(* IEC 61131-3 sources: codesys-api/examples/mqtt_large_payload/st/bcnf_style, 5 files *)

(* ---- AppendGroupBool.st ---- *)
FUNCTION AppendGroupBool : BOOL
// Appends ", 0" or ", 1" to a BCNF-style group line, like INT_TO_STRING(BOOL_TO_INT(x)) in BCNF.
VAR_INPUT
	pBuffer : POINTER TO BYTE;
	Capacity : UDINT;
	Value : BOOL;
END_VAR
VAR_IN_OUT
	Used : UDINT;
END_VAR
// ---- implementation ----
AppendGroupBool := AppendText(pBuffer := pBuffer, Capacity := Capacity, Text := SEL(Value, ', 0', ', 1'), Used := Used);

(* ---- AppendGroupReal.st ---- *)
FUNCTION AppendGroupReal : BOOL
// Appends ", <value>" to a BCNF-style group line, rounded to two decimals exactly as
// FB_InterlockMatrix.StringPublication does. FALSE (and nothing appended) if it would not fit.
VAR_INPUT
	pBuffer : POINTER TO BYTE;
	Capacity : UDINT;
	Value : REAL;
END_VAR
VAR_IN_OUT
	Used : UDINT;
END_VAR
VAR
	Text : STRING(40);
END_VAR
// ---- implementation ----
Text := CONCAT(', ', REAL_TO_STRING(DINT_TO_REAL(TRUNC(Value * 100.0 + SEL(Value >= 0.0, -0.5, 0.5))) / 100.0));
AppendGroupReal := AppendText(pBuffer := pBuffer, Capacity := Capacity, Text := Text, Used := Used);

(* ---- AppendTagLine.st ---- *)
FUNCTION AppendTagLine : BOOL
// Appends "<Name>:<Value>\n", the line format the bridge ingests directly, without a publish map.
// All or nothing: if the whole line doesn't fit, the buffer is left as it was and FALSE is returned.
VAR_INPUT
	pBuffer : POINTER TO BYTE;
	Capacity : UDINT;
	Name : STRING(64);                  // the bridge's tag key for this value
	Value : STRING(40);                 // already formatted, e.g. by REAL_TO_STRING
END_VAR
VAR_IN_OUT
	Used : UDINT;
END_VAR
VAR
	Start : UDINT;
END_VAR
// ---- implementation ----
Start := Used;
AppendTagLine := AppendText(pBuffer := pBuffer, Capacity := Capacity, Text := Name, Used := Used)
	AND_THEN AppendText(pBuffer := pBuffer, Capacity := Capacity, Text := ':', Used := Used)
	AND_THEN AppendText(pBuffer := pBuffer, Capacity := Capacity, Text := Value, Used := Used)
	AND_THEN AppendText(pBuffer := pBuffer, Capacity := Capacity, Text := '$N', Used := Used);
IF NOT AppendTagLine AND pBuffer <> 0 THEN
	Used := Start;
	pBuffer[Start] := 0;
END_IF

(* ---- BcnfPayloadExample.st ---- *)
PROGRAM BcnfPayloadExample
// Sketch of BCNF's StringPublication without the 255-character cap: every group goes into one
// buffer, one "[GROUP, v1, v2, ...]" line per group, so a single publisher sends all of them.
// The values are copied into arrays first; that snapshot is also what a separate MQTT task needs.
// Compiled against the demo project; not run on a PLC.
VAR_INPUT
	IsBuildRequested : BOOL;            // set by the publish timer, not every scan
END_VAR
VAR_OUTPUT
	IsBuildOk : BOOL;                   // FALSE: buffer too small, do not publish this message
	PayloadLength : UDINT;
END_VAR
VAR
	Analog : ARRAY[1..14] OF REAL;      // AIT_1508_V, FIT_1506_F, ... in publish-map order
	Digital : ARRAY[1..9] OF BOOL;      // BCNF_H_E_STOP, LSL_1503_S, ...
	Payload : STRING(4000);
	Used : UDINT;
	Index : INT;
END_VAR
// ---- implementation ----
IF NOT IsBuildRequested THEN
	RETURN;   // BCNF rebuilds its strings every scan today; once per publish is enough
END_IF

// Snapshot (in BCNF: Analog[1] := AIT_1508_V; Analog[2] := FIT_1506_F; ...)

Used := 0;
Payload := '';
IsBuildOk := AppendText(pBuffer := ADR(Payload), Capacity := SIZEOF(Payload), Text := '[BCNF_ANALOG', Used := Used);
FOR Index := 1 TO 14 DO
	IsBuildOk := IsBuildOk AND_THEN AppendGroupReal(pBuffer := ADR(Payload), Capacity := SIZEOF(Payload), Value := Analog[Index], Used := Used);
END_FOR
IsBuildOk := IsBuildOk AND_THEN AppendText(pBuffer := ADR(Payload), Capacity := SIZEOF(Payload), Text := ']$N[BCNF_DIGITAL', Used := Used);
FOR Index := 1 TO 9 DO
	IsBuildOk := IsBuildOk AND_THEN AppendGroupBool(pBuffer := ADR(Payload), Capacity := SIZEOF(Payload), Value := Digital[Index], Used := Used);
END_FOR
IsBuildOk := IsBuildOk AND_THEN AppendText(pBuffer := ADR(Payload), Capacity := SIZEOF(Payload), Text := ']$N', Used := Used);
// ... the same for BCNF_ALARM, BCNF_SETPOINT_1 and _2 (one line once the bridge's publish map
// has a single setpoint entry), BCNF_OUTPUT_OTHER and BCNF_STATUS_STRING.
PayloadLength := Used;
// Publish with PayloadString := ADR(Payload) only when IsBuildOk is TRUE.

(* ---- BcnfStringPublicationCopy.st ---- *)
PROGRAM BcnfStringPublicationCopy
// BCNF's FB_InterlockMatrix.StringPublication, copied verbatim from PLC_BCNF_4_16_26.project, with the
// tags it reads declared using their BCNF types and non-zero values. Generated by
// make_bcnf_copy.py. PLC_PRG calls it every scan when IsBcnfEveryScanEnabled is TRUE,
// to measure what rebuilding BCNF's payload strings every scan costs. Its BuildTagValue action
// builds the same values in the bridge's tag:value line format instead.
VAR
	BCNF_ANALOG_STRING : STRING(255);
	AIT_1508_V : REAL := 16.88;
	FIT_1506_F : REAL := 30.59;
	FIT_1520_F : REAL := 44.30;
	PT_1513_P : REAL := 58.01;
	PT_1516_P : REAL := 71.72;
	QIT_1507_V : REAL := 85.43;
	QIT_1518_V : REAL := 99.14;
	REC_1525_V : REAL := 112.85;
	REJ_1526_V : REAL := 126.56;
	TT_1509_T : REAL := 140.27;
	VFD_1512C_V : REAL := 153.98;
	VFD_1512F_V : REAL := 167.69;
	VFD_1512T_V : REAL := 181.40;
	VFD_1512V_V : REAL := 195.11;
	BCNF_DIGITAL_STRING : STRING(255);
	BCNF_H_E_STOP : BOOL;
	LSL_1503_S : BOOL;
	LSS_E_STOP : BOOL := TRUE;
	LS_1521_S : BOOL;
	LS_1522_S : BOOL;
	LS_1523_S : BOOL := TRUE;
	LS_1524_S : BOOL;
	P_1502FB : BOOL;
	P_1504 : BOOL := TRUE;
	BCNF_ALARM_STRING : STRING(255);
	AIT_1508H : BOOL;
	AIT_1508HH : BOOL;
	AIT_1508L : BOOL := TRUE;
	AIT_1508LL : BOOL;
	BCNF_E_STOP : BOOL;
	BCNF_E_STOPH : BOOL := TRUE;
	BCNF_H_E_STOPH : BOOL;
	CONC_BCNF_PLC_STATUSH : BOOL;
	FIT_1506H : BOOL := TRUE;
	FIT_1506HH : BOOL;
	FIT_1520H : BOOL;
	FIT_1520HH : BOOL := TRUE;
	LSL_1503LL : BOOL;
	LSS_E_STOPH : BOOL;
	LS_1521LL : BOOL := TRUE;
	LS_1522L : BOOL;
	LS_1523H : BOOL;
	LS_1524HH : BOOL := TRUE;
	PT_1513H : BOOL;
	PT_1513HH : BOOL;
	PT_1513L : BOOL := TRUE;
	PT_1513LL : BOOL;
	PT_1516H : BOOL;
	PT_1516HH : BOOL := TRUE;
	PT_1516L : BOOL;
	PT_1516LL : BOOL;
	P_1502FBHH : BOOL := TRUE;
	QIT_1507H : BOOL;
	QIT_1507HH : BOOL;
	QIT_1518H : BOOL := TRUE;
	QIT_1518HH : BOOL;
	TT_1509H : BOOL;
	TT_1509HH : BOOL := TRUE;
	TT_1509L : BOOL;
	TT_1509LL : BOOL;
	VFD_1512CH : BOOL := TRUE;
	VFD_1512CHH : BOOL;
	VFD_1512FH : BOOL;
	VFD_1512FHH : BOOL := TRUE;
	VFD_1512TH : BOOL;
	VFD_1512THH : BOOL;
	VFD_1512VH : BOOL := TRUE;
	VFD_1512VHH : BOOL;
	BCNF_SETPOINT_STRING_1 : STRING(255);
	AIT_1508_HH_SP : REAL := 208.82;
	AIT_1508_H_SP : REAL := 222.53;
	AIT_1508_LL_SP : REAL := 236.24;
	AIT_1508_L_SP : REAL := 249.95;
	FIT_1506_HH_SP : REAL := 263.66;
	FIT_1506_H_SP : REAL := 277.37;
	FIT_1520_HH_SP : REAL := 291.08;
	FIT_1520_H_SP : REAL := 304.79;
	PT_1513_HH_SP : REAL := 318.50;
	PT_1513_H_SP : REAL := 332.21;
	PT_1513_LL_SP : REAL := 345.92;
	PT_1513_L_SP : REAL := 359.63;
	PT_1516_HH_SP : REAL := 373.34;
	PT_1516_H_SP : REAL := 387.05;
	PT_1516_LL_SP : REAL := 400.76;
	PT_1516_L_SP : REAL := 414.47;
	QIT_1507_HH_SP : REAL := 428.18;
	QIT_1507_H_SP : REAL := 441.89;
	QIT_1518_HH_SP : REAL := 455.60;
	QIT_1518_H_SP : REAL := 469.31;
	TT_1509_HH_SP : REAL := 483.02;
	TT_1509_H_SP : REAL := 496.73;
	TT_1509_LL_SP : REAL := 510.44;
	TT_1509_L_SP : REAL := 524.15;
	VFD_1512C_HH_SP : REAL := 537.86;
	VFD_1512C_H_SP : REAL := 551.57;
	BCNF_SETPOINT_STRING_2 : STRING(255);
	VFD_1512F_HH_SP : REAL := 565.28;
	VFD_1512F_H_SP : REAL := 578.99;
	VFD_1512T_HH_SP : REAL := 592.70;
	VFD_1512T_H_SP : REAL := 606.41;
	VFD_1512V_HH_SP : REAL := 620.12;
	VFD_1512V_H_SP : REAL := 633.83;
	BCNF_OUTPUT_OTHER_STRING : STRING(255);
	P_1502_OUTPUT : BOOL;
	VFD_1512FSP : REAL := 647.54;
	VFD_1512SP : REAL := 661.25;
	BCNF_STATUS_STRING : STRING(255);
	Heartbeat : DINT := 18234;
	CONC_BCNF_PLC_STATUS : BOOL := TRUE;
	fullPayload_BCNF_ANALOG_STRING : STRING(255);
	fullPayload_BCNF_DIGITAL_STRING : STRING(255);
	fullPayload_BCNF_ALARM_STRING : STRING(255);
	fullPayload_BCNF_SETPOINT_STRING_1 : STRING(255);
	fullPayload_BCNF_SETPOINT_STRING_2 : STRING(255);
	fullPayload_BCNF_OUTPUT_OTHER_STRING : STRING(255);
	fullPayload_BCNF_STATUS_STRING : STRING(255);
	// BuildTagValue action: the same values as one tag:value line each
	TagValuePayload : STRING(4000);
	TagValueUsed : UDINT;
	IsTagValueBuildOk : BOOL;
END_VAR
// ---- implementation ----
// ===== DATA PUBLICATION STRING BUILDING =====
// This code should be placed in a StringPublication action

// Build BCNF_ANALOG string
BCNF_ANALOG_STRING := '[BCNF_ANALOG, ';
BCNF_ANALOG_STRING := CONCAT(BCNF_ANALOG_STRING, REAL_TO_STRING(DINT_TO_REAL(TRUNC(AIT_1508_V * 100.0 + SEL(AIT_1508_V >= 0.0, -0.5, 0.5))) / 100.0));
BCNF_ANALOG_STRING := CONCAT(BCNF_ANALOG_STRING, ', ');
BCNF_ANALOG_STRING := CONCAT(BCNF_ANALOG_STRING, REAL_TO_STRING(DINT_TO_REAL(TRUNC(FIT_1506_F * 100.0 + SEL(FIT_1506_F >= 0.0, -0.5, 0.5))) / 100.0));
BCNF_ANALOG_STRING := CONCAT(BCNF_ANALOG_STRING, ', ');
BCNF_ANALOG_STRING := CONCAT(BCNF_ANALOG_STRING, REAL_TO_STRING(DINT_TO_REAL(TRUNC(FIT_1520_F * 100.0 + SEL(FIT_1520_F >= 0.0, -0.5, 0.5))) / 100.0));
BCNF_ANALOG_STRING := CONCAT(BCNF_ANALOG_STRING, ', ');
BCNF_ANALOG_STRING := CONCAT(BCNF_ANALOG_STRING, REAL_TO_STRING(DINT_TO_REAL(TRUNC(PT_1513_P * 100.0 + SEL(PT_1513_P >= 0.0, -0.5, 0.5))) / 100.0));
BCNF_ANALOG_STRING := CONCAT(BCNF_ANALOG_STRING, ', ');
BCNF_ANALOG_STRING := CONCAT(BCNF_ANALOG_STRING, REAL_TO_STRING(DINT_TO_REAL(TRUNC(PT_1516_P * 100.0 + SEL(PT_1516_P >= 0.0, -0.5, 0.5))) / 100.0));
BCNF_ANALOG_STRING := CONCAT(BCNF_ANALOG_STRING, ', ');
BCNF_ANALOG_STRING := CONCAT(BCNF_ANALOG_STRING, REAL_TO_STRING(DINT_TO_REAL(TRUNC(QIT_1507_V * 100.0 + SEL(QIT_1507_V >= 0.0, -0.5, 0.5))) / 100.0));
BCNF_ANALOG_STRING := CONCAT(BCNF_ANALOG_STRING, ', ');
BCNF_ANALOG_STRING := CONCAT(BCNF_ANALOG_STRING, REAL_TO_STRING(DINT_TO_REAL(TRUNC(QIT_1518_V * 100.0 + SEL(QIT_1518_V >= 0.0, -0.5, 0.5))) / 100.0));
BCNF_ANALOG_STRING := CONCAT(BCNF_ANALOG_STRING, ', ');
BCNF_ANALOG_STRING := CONCAT(BCNF_ANALOG_STRING, REAL_TO_STRING(DINT_TO_REAL(TRUNC(REC_1525_V * 100.0 + SEL(REC_1525_V >= 0.0, -0.5, 0.5))) / 100.0));
BCNF_ANALOG_STRING := CONCAT(BCNF_ANALOG_STRING, ', ');
BCNF_ANALOG_STRING := CONCAT(BCNF_ANALOG_STRING, REAL_TO_STRING(DINT_TO_REAL(TRUNC(REJ_1526_V * 100.0 + SEL(REJ_1526_V >= 0.0, -0.5, 0.5))) / 100.0));
BCNF_ANALOG_STRING := CONCAT(BCNF_ANALOG_STRING, ', ');
BCNF_ANALOG_STRING := CONCAT(BCNF_ANALOG_STRING, REAL_TO_STRING(DINT_TO_REAL(TRUNC(TT_1509_T * 100.0 + SEL(TT_1509_T >= 0.0, -0.5, 0.5))) / 100.0));
BCNF_ANALOG_STRING := CONCAT(BCNF_ANALOG_STRING, ', ');
BCNF_ANALOG_STRING := CONCAT(BCNF_ANALOG_STRING, REAL_TO_STRING(DINT_TO_REAL(TRUNC(VFD_1512C_V * 100.0 + SEL(VFD_1512C_V >= 0.0, -0.5, 0.5))) / 100.0));
BCNF_ANALOG_STRING := CONCAT(BCNF_ANALOG_STRING, ', ');
BCNF_ANALOG_STRING := CONCAT(BCNF_ANALOG_STRING, REAL_TO_STRING(DINT_TO_REAL(TRUNC(VFD_1512F_V * 100.0 + SEL(VFD_1512F_V >= 0.0, -0.5, 0.5))) / 100.0));
BCNF_ANALOG_STRING := CONCAT(BCNF_ANALOG_STRING, ', ');
BCNF_ANALOG_STRING := CONCAT(BCNF_ANALOG_STRING, REAL_TO_STRING(DINT_TO_REAL(TRUNC(VFD_1512T_V * 100.0 + SEL(VFD_1512T_V >= 0.0, -0.5, 0.5))) / 100.0));
BCNF_ANALOG_STRING := CONCAT(BCNF_ANALOG_STRING, ', ');
BCNF_ANALOG_STRING := CONCAT(BCNF_ANALOG_STRING, REAL_TO_STRING(DINT_TO_REAL(TRUNC(VFD_1512V_V * 100.0 + SEL(VFD_1512V_V >= 0.0, -0.5, 0.5))) / 100.0));
BCNF_ANALOG_STRING := CONCAT(BCNF_ANALOG_STRING, ']');

// Build BCNF_DIGITAL string
BCNF_DIGITAL_STRING := '[BCNF_DIGITAL, ';
BCNF_DIGITAL_STRING := CONCAT(BCNF_DIGITAL_STRING, INT_TO_STRING(BOOL_TO_INT(BCNF_H_E_STOP)));
BCNF_DIGITAL_STRING := CONCAT(BCNF_DIGITAL_STRING, ', ');
BCNF_DIGITAL_STRING := CONCAT(BCNF_DIGITAL_STRING, INT_TO_STRING(BOOL_TO_INT(LSL_1503_S)));
BCNF_DIGITAL_STRING := CONCAT(BCNF_DIGITAL_STRING, ', ');
BCNF_DIGITAL_STRING := CONCAT(BCNF_DIGITAL_STRING, INT_TO_STRING(BOOL_TO_INT(LSS_E_STOP)));
BCNF_DIGITAL_STRING := CONCAT(BCNF_DIGITAL_STRING, ', ');
BCNF_DIGITAL_STRING := CONCAT(BCNF_DIGITAL_STRING, INT_TO_STRING(BOOL_TO_INT(LS_1521_S)));
BCNF_DIGITAL_STRING := CONCAT(BCNF_DIGITAL_STRING, ', ');
BCNF_DIGITAL_STRING := CONCAT(BCNF_DIGITAL_STRING, INT_TO_STRING(BOOL_TO_INT(LS_1522_S)));
BCNF_DIGITAL_STRING := CONCAT(BCNF_DIGITAL_STRING, ', ');
BCNF_DIGITAL_STRING := CONCAT(BCNF_DIGITAL_STRING, INT_TO_STRING(BOOL_TO_INT(LS_1523_S)));
BCNF_DIGITAL_STRING := CONCAT(BCNF_DIGITAL_STRING, ', ');
BCNF_DIGITAL_STRING := CONCAT(BCNF_DIGITAL_STRING, INT_TO_STRING(BOOL_TO_INT(LS_1524_S)));
BCNF_DIGITAL_STRING := CONCAT(BCNF_DIGITAL_STRING, ', ');
BCNF_DIGITAL_STRING := CONCAT(BCNF_DIGITAL_STRING, INT_TO_STRING(BOOL_TO_INT(P_1502FB)));
BCNF_DIGITAL_STRING := CONCAT(BCNF_DIGITAL_STRING, ', ');
BCNF_DIGITAL_STRING := CONCAT(BCNF_DIGITAL_STRING, INT_TO_STRING(BOOL_TO_INT(P_1504)));
BCNF_DIGITAL_STRING := CONCAT(BCNF_DIGITAL_STRING, ']');

// Build BCNF_ALARM string
BCNF_ALARM_STRING := '[BCNF_ALARM, ';
BCNF_ALARM_STRING := CONCAT(BCNF_ALARM_STRING, INT_TO_STRING(BOOL_TO_INT(AIT_1508H)));
BCNF_ALARM_STRING := CONCAT(BCNF_ALARM_STRING, ', ');
BCNF_ALARM_STRING := CONCAT(BCNF_ALARM_STRING, INT_TO_STRING(BOOL_TO_INT(AIT_1508HH)));
BCNF_ALARM_STRING := CONCAT(BCNF_ALARM_STRING, ', ');
BCNF_ALARM_STRING := CONCAT(BCNF_ALARM_STRING, INT_TO_STRING(BOOL_TO_INT(AIT_1508L)));
BCNF_ALARM_STRING := CONCAT(BCNF_ALARM_STRING, ', ');
BCNF_ALARM_STRING := CONCAT(BCNF_ALARM_STRING, INT_TO_STRING(BOOL_TO_INT(AIT_1508LL)));
BCNF_ALARM_STRING := CONCAT(BCNF_ALARM_STRING, ', ');
BCNF_ALARM_STRING := CONCAT(BCNF_ALARM_STRING, INT_TO_STRING(BOOL_TO_INT(BCNF_E_STOP)));
BCNF_ALARM_STRING := CONCAT(BCNF_ALARM_STRING, ', ');
BCNF_ALARM_STRING := CONCAT(BCNF_ALARM_STRING, INT_TO_STRING(BOOL_TO_INT(BCNF_E_STOPH)));
BCNF_ALARM_STRING := CONCAT(BCNF_ALARM_STRING, ', ');
BCNF_ALARM_STRING := CONCAT(BCNF_ALARM_STRING, INT_TO_STRING(BOOL_TO_INT(BCNF_H_E_STOPH)));
BCNF_ALARM_STRING := CONCAT(BCNF_ALARM_STRING, ', ');
BCNF_ALARM_STRING := CONCAT(BCNF_ALARM_STRING, INT_TO_STRING(BOOL_TO_INT(CONC_BCNF_PLC_STATUSH)));
BCNF_ALARM_STRING := CONCAT(BCNF_ALARM_STRING, ', ');
BCNF_ALARM_STRING := CONCAT(BCNF_ALARM_STRING, INT_TO_STRING(BOOL_TO_INT(FIT_1506H)));
BCNF_ALARM_STRING := CONCAT(BCNF_ALARM_STRING, ', ');
BCNF_ALARM_STRING := CONCAT(BCNF_ALARM_STRING, INT_TO_STRING(BOOL_TO_INT(FIT_1506HH)));
BCNF_ALARM_STRING := CONCAT(BCNF_ALARM_STRING, ', ');
BCNF_ALARM_STRING := CONCAT(BCNF_ALARM_STRING, INT_TO_STRING(BOOL_TO_INT(FIT_1520H)));
BCNF_ALARM_STRING := CONCAT(BCNF_ALARM_STRING, ', ');
BCNF_ALARM_STRING := CONCAT(BCNF_ALARM_STRING, INT_TO_STRING(BOOL_TO_INT(FIT_1520HH)));
BCNF_ALARM_STRING := CONCAT(BCNF_ALARM_STRING, ', ');
BCNF_ALARM_STRING := CONCAT(BCNF_ALARM_STRING, INT_TO_STRING(BOOL_TO_INT(LSL_1503LL)));
BCNF_ALARM_STRING := CONCAT(BCNF_ALARM_STRING, ', ');
BCNF_ALARM_STRING := CONCAT(BCNF_ALARM_STRING, INT_TO_STRING(BOOL_TO_INT(LSS_E_STOPH)));
BCNF_ALARM_STRING := CONCAT(BCNF_ALARM_STRING, ', ');
BCNF_ALARM_STRING := CONCAT(BCNF_ALARM_STRING, INT_TO_STRING(BOOL_TO_INT(LS_1521LL)));
BCNF_ALARM_STRING := CONCAT(BCNF_ALARM_STRING, ', ');
BCNF_ALARM_STRING := CONCAT(BCNF_ALARM_STRING, INT_TO_STRING(BOOL_TO_INT(LS_1522L)));
BCNF_ALARM_STRING := CONCAT(BCNF_ALARM_STRING, ', ');
BCNF_ALARM_STRING := CONCAT(BCNF_ALARM_STRING, INT_TO_STRING(BOOL_TO_INT(LS_1523H)));
BCNF_ALARM_STRING := CONCAT(BCNF_ALARM_STRING, ', ');
BCNF_ALARM_STRING := CONCAT(BCNF_ALARM_STRING, INT_TO_STRING(BOOL_TO_INT(LS_1524HH)));
BCNF_ALARM_STRING := CONCAT(BCNF_ALARM_STRING, ', ');
BCNF_ALARM_STRING := CONCAT(BCNF_ALARM_STRING, INT_TO_STRING(BOOL_TO_INT(PT_1513H)));
BCNF_ALARM_STRING := CONCAT(BCNF_ALARM_STRING, ', ');
BCNF_ALARM_STRING := CONCAT(BCNF_ALARM_STRING, INT_TO_STRING(BOOL_TO_INT(PT_1513HH)));
BCNF_ALARM_STRING := CONCAT(BCNF_ALARM_STRING, ', ');
BCNF_ALARM_STRING := CONCAT(BCNF_ALARM_STRING, INT_TO_STRING(BOOL_TO_INT(PT_1513L)));
BCNF_ALARM_STRING := CONCAT(BCNF_ALARM_STRING, ', ');
BCNF_ALARM_STRING := CONCAT(BCNF_ALARM_STRING, INT_TO_STRING(BOOL_TO_INT(PT_1513LL)));
BCNF_ALARM_STRING := CONCAT(BCNF_ALARM_STRING, ', ');
BCNF_ALARM_STRING := CONCAT(BCNF_ALARM_STRING, INT_TO_STRING(BOOL_TO_INT(PT_1516H)));
BCNF_ALARM_STRING := CONCAT(BCNF_ALARM_STRING, ', ');
BCNF_ALARM_STRING := CONCAT(BCNF_ALARM_STRING, INT_TO_STRING(BOOL_TO_INT(PT_1516HH)));
BCNF_ALARM_STRING := CONCAT(BCNF_ALARM_STRING, ', ');
BCNF_ALARM_STRING := CONCAT(BCNF_ALARM_STRING, INT_TO_STRING(BOOL_TO_INT(PT_1516L)));
BCNF_ALARM_STRING := CONCAT(BCNF_ALARM_STRING, ', ');
BCNF_ALARM_STRING := CONCAT(BCNF_ALARM_STRING, INT_TO_STRING(BOOL_TO_INT(PT_1516LL)));
BCNF_ALARM_STRING := CONCAT(BCNF_ALARM_STRING, ', ');
BCNF_ALARM_STRING := CONCAT(BCNF_ALARM_STRING, INT_TO_STRING(BOOL_TO_INT(P_1502FBHH)));
BCNF_ALARM_STRING := CONCAT(BCNF_ALARM_STRING, ', ');
BCNF_ALARM_STRING := CONCAT(BCNF_ALARM_STRING, INT_TO_STRING(BOOL_TO_INT(QIT_1507H)));
BCNF_ALARM_STRING := CONCAT(BCNF_ALARM_STRING, ', ');
BCNF_ALARM_STRING := CONCAT(BCNF_ALARM_STRING, INT_TO_STRING(BOOL_TO_INT(QIT_1507HH)));
BCNF_ALARM_STRING := CONCAT(BCNF_ALARM_STRING, ', ');
BCNF_ALARM_STRING := CONCAT(BCNF_ALARM_STRING, INT_TO_STRING(BOOL_TO_INT(QIT_1518H)));
BCNF_ALARM_STRING := CONCAT(BCNF_ALARM_STRING, ', ');
BCNF_ALARM_STRING := CONCAT(BCNF_ALARM_STRING, INT_TO_STRING(BOOL_TO_INT(QIT_1518HH)));
BCNF_ALARM_STRING := CONCAT(BCNF_ALARM_STRING, ', ');
BCNF_ALARM_STRING := CONCAT(BCNF_ALARM_STRING, INT_TO_STRING(BOOL_TO_INT(TT_1509H)));
BCNF_ALARM_STRING := CONCAT(BCNF_ALARM_STRING, ', ');
BCNF_ALARM_STRING := CONCAT(BCNF_ALARM_STRING, INT_TO_STRING(BOOL_TO_INT(TT_1509HH)));
BCNF_ALARM_STRING := CONCAT(BCNF_ALARM_STRING, ', ');
BCNF_ALARM_STRING := CONCAT(BCNF_ALARM_STRING, INT_TO_STRING(BOOL_TO_INT(TT_1509L)));
BCNF_ALARM_STRING := CONCAT(BCNF_ALARM_STRING, ', ');
BCNF_ALARM_STRING := CONCAT(BCNF_ALARM_STRING, INT_TO_STRING(BOOL_TO_INT(TT_1509LL)));
BCNF_ALARM_STRING := CONCAT(BCNF_ALARM_STRING, ', ');
BCNF_ALARM_STRING := CONCAT(BCNF_ALARM_STRING, INT_TO_STRING(BOOL_TO_INT(VFD_1512CH)));
BCNF_ALARM_STRING := CONCAT(BCNF_ALARM_STRING, ', ');
BCNF_ALARM_STRING := CONCAT(BCNF_ALARM_STRING, INT_TO_STRING(BOOL_TO_INT(VFD_1512CHH)));
BCNF_ALARM_STRING := CONCAT(BCNF_ALARM_STRING, ', ');
BCNF_ALARM_STRING := CONCAT(BCNF_ALARM_STRING, INT_TO_STRING(BOOL_TO_INT(VFD_1512FH)));
BCNF_ALARM_STRING := CONCAT(BCNF_ALARM_STRING, ', ');
BCNF_ALARM_STRING := CONCAT(BCNF_ALARM_STRING, INT_TO_STRING(BOOL_TO_INT(VFD_1512FHH)));
BCNF_ALARM_STRING := CONCAT(BCNF_ALARM_STRING, ', ');
BCNF_ALARM_STRING := CONCAT(BCNF_ALARM_STRING, INT_TO_STRING(BOOL_TO_INT(VFD_1512TH)));
BCNF_ALARM_STRING := CONCAT(BCNF_ALARM_STRING, ', ');
BCNF_ALARM_STRING := CONCAT(BCNF_ALARM_STRING, INT_TO_STRING(BOOL_TO_INT(VFD_1512THH)));
BCNF_ALARM_STRING := CONCAT(BCNF_ALARM_STRING, ', ');
BCNF_ALARM_STRING := CONCAT(BCNF_ALARM_STRING, INT_TO_STRING(BOOL_TO_INT(VFD_1512VH)));
BCNF_ALARM_STRING := CONCAT(BCNF_ALARM_STRING, ', ');
BCNF_ALARM_STRING := CONCAT(BCNF_ALARM_STRING, INT_TO_STRING(BOOL_TO_INT(VFD_1512VHH)));
BCNF_ALARM_STRING := CONCAT(BCNF_ALARM_STRING, ']');

// Build BCNF_SETPOINT string part 1
BCNF_SETPOINT_STRING_1 := '[BCNF_SETPOINT_1, ';
BCNF_SETPOINT_STRING_1 := CONCAT(BCNF_SETPOINT_STRING_1, REAL_TO_STRING(DINT_TO_REAL(TRUNC(AIT_1508_HH_SP * 100.0 + SEL(AIT_1508_HH_SP >= 0.0, -0.5, 0.5))) / 100.0));
BCNF_SETPOINT_STRING_1 := CONCAT(BCNF_SETPOINT_STRING_1, ', ');
BCNF_SETPOINT_STRING_1 := CONCAT(BCNF_SETPOINT_STRING_1, REAL_TO_STRING(DINT_TO_REAL(TRUNC(AIT_1508_H_SP * 100.0 + SEL(AIT_1508_H_SP >= 0.0, -0.5, 0.5))) / 100.0));
BCNF_SETPOINT_STRING_1 := CONCAT(BCNF_SETPOINT_STRING_1, ', ');
BCNF_SETPOINT_STRING_1 := CONCAT(BCNF_SETPOINT_STRING_1, REAL_TO_STRING(DINT_TO_REAL(TRUNC(AIT_1508_LL_SP * 100.0 + SEL(AIT_1508_LL_SP >= 0.0, -0.5, 0.5))) / 100.0));
BCNF_SETPOINT_STRING_1 := CONCAT(BCNF_SETPOINT_STRING_1, ', ');
BCNF_SETPOINT_STRING_1 := CONCAT(BCNF_SETPOINT_STRING_1, REAL_TO_STRING(DINT_TO_REAL(TRUNC(AIT_1508_L_SP * 100.0 + SEL(AIT_1508_L_SP >= 0.0, -0.5, 0.5))) / 100.0));
BCNF_SETPOINT_STRING_1 := CONCAT(BCNF_SETPOINT_STRING_1, ', ');
BCNF_SETPOINT_STRING_1 := CONCAT(BCNF_SETPOINT_STRING_1, REAL_TO_STRING(DINT_TO_REAL(TRUNC(FIT_1506_HH_SP * 100.0 + SEL(FIT_1506_HH_SP >= 0.0, -0.5, 0.5))) / 100.0));
BCNF_SETPOINT_STRING_1 := CONCAT(BCNF_SETPOINT_STRING_1, ', ');
BCNF_SETPOINT_STRING_1 := CONCAT(BCNF_SETPOINT_STRING_1, REAL_TO_STRING(DINT_TO_REAL(TRUNC(FIT_1506_H_SP * 100.0 + SEL(FIT_1506_H_SP >= 0.0, -0.5, 0.5))) / 100.0));
BCNF_SETPOINT_STRING_1 := CONCAT(BCNF_SETPOINT_STRING_1, ', ');
BCNF_SETPOINT_STRING_1 := CONCAT(BCNF_SETPOINT_STRING_1, REAL_TO_STRING(DINT_TO_REAL(TRUNC(FIT_1520_HH_SP * 100.0 + SEL(FIT_1520_HH_SP >= 0.0, -0.5, 0.5))) / 100.0));
BCNF_SETPOINT_STRING_1 := CONCAT(BCNF_SETPOINT_STRING_1, ', ');
BCNF_SETPOINT_STRING_1 := CONCAT(BCNF_SETPOINT_STRING_1, REAL_TO_STRING(DINT_TO_REAL(TRUNC(FIT_1520_H_SP * 100.0 + SEL(FIT_1520_H_SP >= 0.0, -0.5, 0.5))) / 100.0));
BCNF_SETPOINT_STRING_1 := CONCAT(BCNF_SETPOINT_STRING_1, ', ');
BCNF_SETPOINT_STRING_1 := CONCAT(BCNF_SETPOINT_STRING_1, REAL_TO_STRING(DINT_TO_REAL(TRUNC(PT_1513_HH_SP * 100.0 + SEL(PT_1513_HH_SP >= 0.0, -0.5, 0.5))) / 100.0));
BCNF_SETPOINT_STRING_1 := CONCAT(BCNF_SETPOINT_STRING_1, ', ');
BCNF_SETPOINT_STRING_1 := CONCAT(BCNF_SETPOINT_STRING_1, REAL_TO_STRING(DINT_TO_REAL(TRUNC(PT_1513_H_SP * 100.0 + SEL(PT_1513_H_SP >= 0.0, -0.5, 0.5))) / 100.0));
BCNF_SETPOINT_STRING_1 := CONCAT(BCNF_SETPOINT_STRING_1, ', ');
BCNF_SETPOINT_STRING_1 := CONCAT(BCNF_SETPOINT_STRING_1, REAL_TO_STRING(DINT_TO_REAL(TRUNC(PT_1513_LL_SP * 100.0 + SEL(PT_1513_LL_SP >= 0.0, -0.5, 0.5))) / 100.0));
BCNF_SETPOINT_STRING_1 := CONCAT(BCNF_SETPOINT_STRING_1, ', ');
BCNF_SETPOINT_STRING_1 := CONCAT(BCNF_SETPOINT_STRING_1, REAL_TO_STRING(DINT_TO_REAL(TRUNC(PT_1513_L_SP * 100.0 + SEL(PT_1513_L_SP >= 0.0, -0.5, 0.5))) / 100.0));
BCNF_SETPOINT_STRING_1 := CONCAT(BCNF_SETPOINT_STRING_1, ', ');
BCNF_SETPOINT_STRING_1 := CONCAT(BCNF_SETPOINT_STRING_1, REAL_TO_STRING(DINT_TO_REAL(TRUNC(PT_1516_HH_SP * 100.0 + SEL(PT_1516_HH_SP >= 0.0, -0.5, 0.5))) / 100.0));
BCNF_SETPOINT_STRING_1 := CONCAT(BCNF_SETPOINT_STRING_1, ', ');
BCNF_SETPOINT_STRING_1 := CONCAT(BCNF_SETPOINT_STRING_1, REAL_TO_STRING(DINT_TO_REAL(TRUNC(PT_1516_H_SP * 100.0 + SEL(PT_1516_H_SP >= 0.0, -0.5, 0.5))) / 100.0));
BCNF_SETPOINT_STRING_1 := CONCAT(BCNF_SETPOINT_STRING_1, ', ');
BCNF_SETPOINT_STRING_1 := CONCAT(BCNF_SETPOINT_STRING_1, REAL_TO_STRING(DINT_TO_REAL(TRUNC(PT_1516_LL_SP * 100.0 + SEL(PT_1516_LL_SP >= 0.0, -0.5, 0.5))) / 100.0));
BCNF_SETPOINT_STRING_1 := CONCAT(BCNF_SETPOINT_STRING_1, ', ');
BCNF_SETPOINT_STRING_1 := CONCAT(BCNF_SETPOINT_STRING_1, REAL_TO_STRING(DINT_TO_REAL(TRUNC(PT_1516_L_SP * 100.0 + SEL(PT_1516_L_SP >= 0.0, -0.5, 0.5))) / 100.0));
BCNF_SETPOINT_STRING_1 := CONCAT(BCNF_SETPOINT_STRING_1, ', ');
BCNF_SETPOINT_STRING_1 := CONCAT(BCNF_SETPOINT_STRING_1, REAL_TO_STRING(DINT_TO_REAL(TRUNC(QIT_1507_HH_SP * 100.0 + SEL(QIT_1507_HH_SP >= 0.0, -0.5, 0.5))) / 100.0));
BCNF_SETPOINT_STRING_1 := CONCAT(BCNF_SETPOINT_STRING_1, ', ');
BCNF_SETPOINT_STRING_1 := CONCAT(BCNF_SETPOINT_STRING_1, REAL_TO_STRING(DINT_TO_REAL(TRUNC(QIT_1507_H_SP * 100.0 + SEL(QIT_1507_H_SP >= 0.0, -0.5, 0.5))) / 100.0));
BCNF_SETPOINT_STRING_1 := CONCAT(BCNF_SETPOINT_STRING_1, ', ');
BCNF_SETPOINT_STRING_1 := CONCAT(BCNF_SETPOINT_STRING_1, REAL_TO_STRING(DINT_TO_REAL(TRUNC(QIT_1518_HH_SP * 100.0 + SEL(QIT_1518_HH_SP >= 0.0, -0.5, 0.5))) / 100.0));
BCNF_SETPOINT_STRING_1 := CONCAT(BCNF_SETPOINT_STRING_1, ', ');
BCNF_SETPOINT_STRING_1 := CONCAT(BCNF_SETPOINT_STRING_1, REAL_TO_STRING(DINT_TO_REAL(TRUNC(QIT_1518_H_SP * 100.0 + SEL(QIT_1518_H_SP >= 0.0, -0.5, 0.5))) / 100.0));
BCNF_SETPOINT_STRING_1 := CONCAT(BCNF_SETPOINT_STRING_1, ', ');
BCNF_SETPOINT_STRING_1 := CONCAT(BCNF_SETPOINT_STRING_1, REAL_TO_STRING(DINT_TO_REAL(TRUNC(TT_1509_HH_SP * 100.0 + SEL(TT_1509_HH_SP >= 0.0, -0.5, 0.5))) / 100.0));
BCNF_SETPOINT_STRING_1 := CONCAT(BCNF_SETPOINT_STRING_1, ', ');
BCNF_SETPOINT_STRING_1 := CONCAT(BCNF_SETPOINT_STRING_1, REAL_TO_STRING(DINT_TO_REAL(TRUNC(TT_1509_H_SP * 100.0 + SEL(TT_1509_H_SP >= 0.0, -0.5, 0.5))) / 100.0));
BCNF_SETPOINT_STRING_1 := CONCAT(BCNF_SETPOINT_STRING_1, ', ');
BCNF_SETPOINT_STRING_1 := CONCAT(BCNF_SETPOINT_STRING_1, REAL_TO_STRING(DINT_TO_REAL(TRUNC(TT_1509_LL_SP * 100.0 + SEL(TT_1509_LL_SP >= 0.0, -0.5, 0.5))) / 100.0));
BCNF_SETPOINT_STRING_1 := CONCAT(BCNF_SETPOINT_STRING_1, ', ');
BCNF_SETPOINT_STRING_1 := CONCAT(BCNF_SETPOINT_STRING_1, REAL_TO_STRING(DINT_TO_REAL(TRUNC(TT_1509_L_SP * 100.0 + SEL(TT_1509_L_SP >= 0.0, -0.5, 0.5))) / 100.0));
BCNF_SETPOINT_STRING_1 := CONCAT(BCNF_SETPOINT_STRING_1, ', ');
BCNF_SETPOINT_STRING_1 := CONCAT(BCNF_SETPOINT_STRING_1, REAL_TO_STRING(DINT_TO_REAL(TRUNC(VFD_1512C_HH_SP * 100.0 + SEL(VFD_1512C_HH_SP >= 0.0, -0.5, 0.5))) / 100.0));
BCNF_SETPOINT_STRING_1 := CONCAT(BCNF_SETPOINT_STRING_1, ', ');
BCNF_SETPOINT_STRING_1 := CONCAT(BCNF_SETPOINT_STRING_1, REAL_TO_STRING(DINT_TO_REAL(TRUNC(VFD_1512C_H_SP * 100.0 + SEL(VFD_1512C_H_SP >= 0.0, -0.5, 0.5))) / 100.0));
BCNF_SETPOINT_STRING_1 := CONCAT(BCNF_SETPOINT_STRING_1, ']');
// Build BCNF_SETPOINT string part 2
BCNF_SETPOINT_STRING_2 := '[BCNF_SETPOINT_2, ';
BCNF_SETPOINT_STRING_2 := CONCAT(BCNF_SETPOINT_STRING_2, REAL_TO_STRING(DINT_TO_REAL(TRUNC(VFD_1512F_HH_SP * 100.0 + SEL(VFD_1512F_HH_SP >= 0.0, -0.5, 0.5))) / 100.0));
BCNF_SETPOINT_STRING_2 := CONCAT(BCNF_SETPOINT_STRING_2, ', ');
BCNF_SETPOINT_STRING_2 := CONCAT(BCNF_SETPOINT_STRING_2, REAL_TO_STRING(DINT_TO_REAL(TRUNC(VFD_1512F_H_SP * 100.0 + SEL(VFD_1512F_H_SP >= 0.0, -0.5, 0.5))) / 100.0));
BCNF_SETPOINT_STRING_2 := CONCAT(BCNF_SETPOINT_STRING_2, ', ');
BCNF_SETPOINT_STRING_2 := CONCAT(BCNF_SETPOINT_STRING_2, REAL_TO_STRING(DINT_TO_REAL(TRUNC(VFD_1512T_HH_SP * 100.0 + SEL(VFD_1512T_HH_SP >= 0.0, -0.5, 0.5))) / 100.0));
BCNF_SETPOINT_STRING_2 := CONCAT(BCNF_SETPOINT_STRING_2, ', ');
BCNF_SETPOINT_STRING_2 := CONCAT(BCNF_SETPOINT_STRING_2, REAL_TO_STRING(DINT_TO_REAL(TRUNC(VFD_1512T_H_SP * 100.0 + SEL(VFD_1512T_H_SP >= 0.0, -0.5, 0.5))) / 100.0));
BCNF_SETPOINT_STRING_2 := CONCAT(BCNF_SETPOINT_STRING_2, ', ');
BCNF_SETPOINT_STRING_2 := CONCAT(BCNF_SETPOINT_STRING_2, REAL_TO_STRING(DINT_TO_REAL(TRUNC(VFD_1512V_HH_SP * 100.0 + SEL(VFD_1512V_HH_SP >= 0.0, -0.5, 0.5))) / 100.0));
BCNF_SETPOINT_STRING_2 := CONCAT(BCNF_SETPOINT_STRING_2, ', ');
BCNF_SETPOINT_STRING_2 := CONCAT(BCNF_SETPOINT_STRING_2, REAL_TO_STRING(DINT_TO_REAL(TRUNC(VFD_1512V_H_SP * 100.0 + SEL(VFD_1512V_H_SP >= 0.0, -0.5, 0.5))) / 100.0));
BCNF_SETPOINT_STRING_2 := CONCAT(BCNF_SETPOINT_STRING_2, ']');

// Build BCNF_OUTPUT_OTHER string
BCNF_OUTPUT_OTHER_STRING := '[BCNF_OUTPUT_OTHER, ';
BCNF_OUTPUT_OTHER_STRING := CONCAT(BCNF_OUTPUT_OTHER_STRING, INT_TO_STRING(BOOL_TO_INT(P_1502_OUTPUT)));
BCNF_OUTPUT_OTHER_STRING := CONCAT(BCNF_OUTPUT_OTHER_STRING, ', ');
BCNF_OUTPUT_OTHER_STRING := CONCAT(BCNF_OUTPUT_OTHER_STRING, REAL_TO_STRING(DINT_TO_REAL(TRUNC(VFD_1512FSP * 100.0 + SEL(VFD_1512FSP >= 0.0, -0.5, 0.5))) / 100.0));
BCNF_OUTPUT_OTHER_STRING := CONCAT(BCNF_OUTPUT_OTHER_STRING, ', ');
BCNF_OUTPUT_OTHER_STRING := CONCAT(BCNF_OUTPUT_OTHER_STRING, REAL_TO_STRING(DINT_TO_REAL(TRUNC(VFD_1512SP * 100.0 + SEL(VFD_1512SP >= 0.0, -0.5, 0.5))) / 100.0));
BCNF_OUTPUT_OTHER_STRING := CONCAT(BCNF_OUTPUT_OTHER_STRING, ']');

// ===== PAYLOAD ASSIGNMENTS =====
// ----- Build Status String -----
// Format: [BCNF_STATUS_STRING, Heartbeat, STATUS]
BCNF_STATUS_STRING := '[BCNF_STATUS_STRING, ';
BCNF_STATUS_STRING := CONCAT(BCNF_STATUS_STRING, DINT_TO_STRING(Heartbeat));
BCNF_STATUS_STRING := CONCAT(BCNF_STATUS_STRING, ', ');
BCNF_STATUS_STRING := CONCAT(BCNF_STATUS_STRING, BOOL_TO_STRING(CONC_BCNF_PLC_STATUS));
BCNF_STATUS_STRING := CONCAT(BCNF_STATUS_STRING, ']');

fullPayload_BCNF_ANALOG_STRING := BCNF_ANALOG_STRING;
fullPayload_BCNF_DIGITAL_STRING := BCNF_DIGITAL_STRING;
fullPayload_BCNF_ALARM_STRING := BCNF_ALARM_STRING;
fullPayload_BCNF_SETPOINT_STRING_1 := BCNF_SETPOINT_STRING_1;
fullPayload_BCNF_SETPOINT_STRING_2 := BCNF_SETPOINT_STRING_2;
fullPayload_BCNF_OUTPUT_OTHER_STRING := BCNF_OUTPUT_OTHER_STRING;
fullPayload_BCNF_STATUS_STRING := BCNF_STATUS_STRING;
